(* IEC 61131-3 sources: JingjiangMoonbox/Application/Application/数据类型/通讯协议/月影, 10 files *)

(* ---- StParam_Mailbox.st ---- *)
(*@CES
Name=StParam_Mailbox
Type=Gvl
TypeGuid=2db5746d-d284-4425-9f7f-2663a34b0ebc
Guid=28298cb9-a045-46a0-b057-5251b4c14df2
HasDeclaration=True
HasImplementation=False
*)
{DECLARATION}
{attribute 'pack_mode' := '1'}
TYPE StParam_Mailbox :
STRUCT
	dwSemaphore						:DWORD;(*通讯旗语						*)
	dwPlateAdjustmentProf			:DWORD;(*纵向版快速调整量/bit24~bit31为请求信号/低24bit用来表示要调整的量<单位:0.01mm>/ 	*)
	iRapidAdjProf_h					:INT  ;(*横向快速对版量描述				*)
	iGateSa							:INT  ;(*第一波门位置					*)
	iGateSaEx						:INT  ;(*第二波门位置					*)
	rAdjust_V						:REAL ;(*纵向版修正量					*)
	rAdjust_H						:REAL ;(*横向版修正量					*)
	dwFlag_Ctl						:DWORD;(*套色控制标志					*)
	dwFlag_Sts						:DWORD;(*套色状态标志					*)
	wButtonFun_Lamp					:WORD ;(*HMI界面按钮及指示灯			*)
	wSwitchFun						:WORD ;(*界面开关*)
	wRsv							:WORD;
//2025.11.7.142851先把数据统一了，dwSlaveBtn_HMI分两个word,一个暂时baoliu
//	dwSlaveBtn_HMI					:DWORD;(*界面按钮						*)
	rStep_Pressure_Prn_Net			:REAL ;(*版辊网辊按钮步进量				*)
	rLong_Step_Roller_Pressure		:REAL ;(*色组压力控制长步进值			*)
	rShort_Step_Roller_Pressure		:REAL ;(*色组压力控制短步进值			*)
	wAirInletWindDoorValue			:WORD ;(*进风口风门开度值				*)
	wAirExhaustWindDoorValue		:WORD ;(*排风口风门开度值				*)
	wAirReturnWindDoorValue			:WORD ;(*回风口风门开度值				*)
	dwCtlBits_UnitBaseCraft			:DWORD;(*界面工艺开关及状态				*)
	wHz_UnitInkRoller_ManuallySet	:WORD ;(*递墨辊手动频率					*)
	wCoeff_UnitInkRoller_Auto		:WORD ;(*递墨辊自动系数					*)
	wHz_UnitScraper_ManuallySet		:WORD ;(*刮刀手动频率					*)
	wCoeff_UnitScraper_Auto			:WORD ;(*刮刀自动系数					*)
	wHz_UnitHotWind					:WORD ;(*热风频率						*)
	wHz_UnitHotWind_2				:WORD ;(*热风2频率						*)
	wSV_UnitTemCtl					:WORD ;(*加热设定温度					*)
	wUnit_output_I					:WORD ;(*IO监控输出1					*)
	wUnit_output_II					:WORD ;(*IO监控输出2					*)
	//xi.hy//新增
	bySignalSelect					:BYTE; (*光纤电眼信号选择*)
	rOffset_T1						:REAL;	//T1路光纤偏移
	rSource_Light_T1       			:REAL;  //T1路光纤光源
	rBias_T1			  			:REAL;  //T1路光纤电眼偏置
	rBrightness_Light_T1			:REAL;  //T1路光纤电眼亮度

	rOffset_T2						:REAL;  //T2路光纤偏移
	rSource_Light_T2				:REAL;  //T2路光纤光源
	rBias_T2						:REAL;  //T2路光纤电眼偏置
	rBrightness_Light_T2			:REAL;  //T2路光纤电眼亮度

	(*2025.8.14.143359增加一些参数*)
// 	wAccButton_Count				: WORD;
// 	wDecButton_Count			: WORD;
// 	wUpAdjButton_Count			: WORD;
// 	wDnAdjButton_Count			: WORD;
// 	wLeftAdjButton_Count			: WORD;
// 	wRightAdjButton_Count			: WORD;
// 	wAlarmButton_Count			: WORD;

	rHz_AxisAirBlowning_ManuallySet			: REAL;
	rHz_AxisAirExhaust_ManuallySet		: REAL;

	wSlaveBtn_HMI		: WORD;    //.0 版辊操作侧靠近
								   //.1 版辊操作侧远离
								   //.2 版辊平行靠近
								   //.3 版辊平行远离
								   //.4 版辊传动侧靠近
								   //.5 版辊传动侧远离
								   //.6 网辊操作侧靠近
								   //.7 网辊操作侧远离
								   //.8 网辊平行靠近
								   //.9 网辊平行远离
								   //.10 网辊传动侧靠近
								   //.11 网辊传动侧远离
								   //.12 版辊标定
								   //.13 网辊标定
								   //.14 张带棍标定
							 	   //.15 版辊合压
	wSlaveBtn_HMI2		: WORD;
									//. 0  版辊离压
									//. 1 网辊合压
									//. 2 网辊离压
									//. 3 版辊换版
									//. 4 网辊换版
									//. 5 自动换版
									//. 6 换版完成
									// .7 显示换版状态
	wButtonAndSwitch_ChaoXu	: WORD;	//.0 匀墨
										//.1 网辊锁轴
										//.2 充气
										//.3 墨盘电磁阀升
										//.4 照明
										//.5 显示是否修改版周
										//.6 确认修改版周
										//.7
										//.8
										//.9 版辊单动
										//.10 底辊单动
										//.11 合压
										//.12 离压
										//.13 横向左移
										//.14 横向右移

	uiRsv_data					: UINT;//压力电机步进量2026.02.07.143804
	iStep_Horz_Use						: INT;

	//xi.hy
	wState_FiberMove:WORD;	//光纤行走状态
						//.0 行走电机运动中
						//.1 基准色位置确认
						//.2 手动左移
						//.3 手动右移
						//.4 定长运动启动使能
						//.5 回零正限位触发
						//.6 宽度计算成功标志
						//.7 电机读取回来的限位信号
						//.8 基准位置同步完成
						//.9 基准位置同步中
						//.10 从站计算宽度使能
						//.11
						//.12
						//.13
						//.14
						//.15
	wAlarm_FiberMove:WORD;		//光纤行走报警
	iFiberMoveDistanceIn:INT;	//光纤行走距离输入 *10
	iPosCur_FiberMove:INT;		//光纤行走当前位置*10
	iWidth_FindMarkCenter:INT;	//光纤行走 计算出来的宽度*100
	//2026.5.9.182337
	//2026.04.28.132649 xi.hy新增@七号开始
	iStsSlave_FiberMove:INT;  // 光纤行走 从站运动状态机
	//2026.05.28.181612
	iFiberMoveBasePosFromSlave:INT;//基准位置@来自从站

END_STRUCT
END_TYPE

{IMPLEMENTATION}

(* ---- StParam_PDU_Dn.st ---- *)
(*@CES
Name=StParam_PDU_Dn
Type=Gvl
TypeGuid=2db5746d-d284-4425-9f7f-2663a34b0ebc
Guid=7cc610ea-6431-4c4c-b72a-07e9312a874d
HasDeclaration=True
HasImplementation=False
*)
{DECLARATION}
{attribute 'pack_mode' := '1'}
TYPE StParam_PDU_Dn :
STRUCT
	byPkgId						: BYTE;(*数据包ID*)
	abyPayLoad					: ARRAY [1..57] OF BYTE;(*数据可变区域*)
	wCHK						: WORD;(*校验码*)
END_STRUCT
END_TYPE

{IMPLEMENTATION}

(* ---- StParam_PDU_Up.st ---- *)
(*@CES
Name=StParam_PDU_Up
Type=Gvl
TypeGuid=2db5746d-d284-4425-9f7f-2663a34b0ebc
Guid=86ab3953-ed0c-4c63-9744-6672adabd60d
HasDeclaration=True
HasImplementation=False
*)
{DECLARATION}
{attribute 'pack_mode' := '1'}
TYPE StParam_PDU_Up :
STRUCT
	byPkgId						: BYTE;(*数据包ID*)
	abyPayLoad					: ARRAY [1..45] OF BYTE;(*数据可变区域*)
	wCHK						: WORD;(*校验码*)
	byIDX_V						: BYTE;(*纵向误差索引*)
	byIDX_H						: BYTE;(* 横向误差索引 *)
	iErr_V_Raw					: INT;(*纵向误差原始值-跟前色*)
	iErr_H_Raw					: INT;(*横向误差原始值-跟前色*)
	iErr_V_Raw_1				: INT;(*纵向误差原始值-跟任意色*)
	iErr_H_Raw_1				: INT;(*横向误差原始值-跟任意色*)
	uiFSampleCounter			: UINT;(*精采样计数*)
END_STRUCT
END_TYPE

{IMPLEMENTATION}

(* ---- StPdu_Dn_91.st ---- *)
(*@CES
Name=StPdu_Dn_91
Type=Gvl
TypeGuid=2db5746d-d284-4425-9f7f-2663a34b0ebc
Guid=22e1e21e-e973-4286-a59d-d3b41682a852
HasDeclaration=True
HasImplementation=False
*)
{DECLARATION}
{attribute 'pack_mode' := '1'}
TYPE StPdu_Dn_91 :
STRUCT
	byUnitId					:BYTE  ;(*机组号+系ID(最高位为系ID)*)
	rGirth_Sam					:REAL  ;(*采样版周长*)
	uiNum_Sam					:WORD  ;(*采样减速比分子*)
	uiDen_Sam					:WORD  ;(*采样减速比分母*)
	byCurrUsrLevel				:BYTE  ;(*用户权限*)
	iCompanyId					:INT   ;(*用户编号*)
	byLanguageId				:BYTE  ;(*语言选择*)
	byMinutes_ScrAutoSleep		:BYTE  ;(*屏幕休眠时间*)
	wUnit_input_I				:WORD  ;(*色组IO输入1*)
	wUnit_input_II				:WORD  ;(*色组IO输入2*)
	wUnit_input_III				:WORD  ;(*色组IO输入3*)
	wVelocity					:WORD  ;(*主机速度，单位0.1m/min*)
	wVel_Axis					:WORD  ;(*轴速度，单位0.1m/min*)
//	wComplexBit					:WORD  ;(*复合控制位描述*)
	wAxis_RollerDn				:WORD  ;(*轴压辊状态(bit0-1U,bit15-16U)*)
	wAxis_Alarm_Prn				:WORD  ;(*色组版辊报警状态(bit0-1U,bit15-16U)*)
	dwAlarmCode					:DWORD ;(*轴报警码*)
	wComplexFlag_AxisInching	:WORD  ;(*所有轴的单运行状态*)
	wComplexFlag_Linkage		:WORD  ;(*所有轴的联动状态*)
	wComplexFlag_Estop			:DWORD ;(*所有轴的急停状态*)
	wHMI_SwitchSts				:WORD  ;(*色组人机界面开关状态*)
	wSts_HorzManuPreReg			:WORD  ;(*横向手动预套准状态*)
	iPos_HorzManuPreReg			:INT   ;(*横向手动预套准位置*)
(*2025.8.6.205703增加*)
	bySts_Flag					:BYTE;(*色组状态*)
(*	dwAxis_SkipTheHeader 		:DWORD;(*让料头标志*)*)
	bySts_Machine				:BYTE;
	(*
		bit0: 印刷标志
		bit1: 空转标志
		bit2:
	*)
	//2025.11.14.155203||把误差状态发到从站，用于从站人机屏保实现9-1=8；
	byErrSts_V					: BYTE;
//用两个预留放低通滤波频率2025.11.15.132130|niu.j|8-2=6
	//Filter原本的wRsv在这里改一下改为从站精采样数据低通滤波频率
	uilowpasscutoff_hz				:UINT;

	abyRsv_91					:ARRAY [1..6] OF BYTE  ;(*预留空间*)
END_STRUCT
END_TYPE

{IMPLEMENTATION}

(* ---- StPdu_Dn_92.st ---- *)
(*@CES
Name=StPdu_Dn_92
Type=Gvl
TypeGuid=2db5746d-d284-4425-9f7f-2663a34b0ebc
Guid=45573361-4128-408d-910f-d2643f065581
HasDeclaration=True
HasImplementation=False
*)
{DECLARATION}
{attribute 'pack_mode' := '1'}
TYPE StPdu_Dn_92 :
STRUCT
	iCurveViewMaxRange				:INT;(*误差曲线量程上限		*)
	bySignalGain					:BYTE;(*光电眼IO控制			*)
	byMarkTypeId					:BYTE;(*标记形式				*)
	byMarkArrangeModalId			:BYTE;(*标记排列形式			*)
	byFakeThreshold_V				:BYTE;(*纵向飞点阀值@丝			*)
	byFakeThreshold_H				:BYTE;(*横向飞点阀值@丝			*)
	rAlarm_V						:REAL;(*纵向报警值@mm			*)
	rAlarm_H						:REAL;(*横向报警值@mm			*)
	byAve_v_extra_V					:BYTE;(*套色误差显示平均次数	*)
	byAve_v_extra_H					:BYTE;(*套色误差显示平均次数	*)
(*	dwFlag_Sts						: DWORD;(* 状态标志 *)
(*												/bit0.纵向自动 *)
(*												/bit1.横向自动
												/bit9.双极性*)
(*												/ *)
*)
	iGateWidthPhy					: INT ;(*波门宽度				*)
	byTriangleMark_SideC			: BYTE;(*梯形标记三角形纵向边长	*)
	byTriangleMark_SideB			: BYTE;(*梯形标记三角形横向边长	*)
	bySysSamplePrecision			: BYTE;(*系统采样精度			*)
	byArcFineSampleType				: BYTE;(*套色采样方式			*)
	iSampleCfgParam_ctl				: INT ;(*采样控制参数里的ctl		*)
	byColorIdCurrent				: BYTE;(*当前色序				*)
	byColorIdFollow					: BYTE;(*跟踪色序				*)
	abyColorIdList					: ARRAY [1..16] OF BYTE;(*色序列表				*)
	//bySignalSelect					:BYTE;(*光纤电眼信号选择		*)
	xEnable_Arc						: BOOL;(*套印使能开关			*)
	uiSource_Light_T1_Cur			: UINT;
	uiSource_Light_T2_Cur			: UINT;

	//xi.hy2026.5.9.104409
	wDirAndMode_FiberMove			:WORD;//光纤行走的方向和模式:低位方向,高位模式：0不运动 1连续运动 2定长运动 3回零运动
	uiVel_FiberMove					:UINT;//光纤行走的速度:mm/s *10
	uiDistanceOut_FiberMove			:UINT;//光纤行走的输出距离:mm *10
	uiPulsePerCycle_FiberMove		:UINT;//光纤行走的单圈脉冲:pluse

	abyRsv_92						: ARRAY [1..1] OF BYTE;(*套色参数预留			*)
END_STRUCT
END_TYPE

{IMPLEMENTATION}

(* ---- StPdu_Dn_93.st ---- *)
(*@CES
Name=StPdu_Dn_93
Type=Gvl
TypeGuid=2db5746d-d284-4425-9f7f-2663a34b0ebc
Guid=1bb7fc47-9e93-466c-a1c5-84993bb7c104
HasDeclaration=True
HasImplementation=False
*)
{DECLARATION}
{attribute 'pack_mode' := '1'}
TYPE StPdu_Dn_93 :
STRUCT
	dwControlComplexBits		:DWORD;(*开关状态			*)
	wHz_UnitInkRoller_CurrWR	:WORD ;(*递墨辊最终写入频率	*)
	wHz_UnitScraper_CurrWR		:WORD ;(*刮刀写入频率		*)
	wHz_UnitHotWind_CurrWR		:WORD ;(*热风写入频率		*)
	wHz_UnitHotWind2_CurrWR		:WORD ;(*热风2写入频率		*)
	rPV_UnitTemCtl				:REAL ;(*当前温度			*)
	wSTS_UnitTemCtl				:WORD ;(*温控状态			*)
(*2025.8.6.212214增加*)
	wHotWind_Print				:WORD;(*热风打开色组号*)
	byDriverType_Hor			:BYTE;(*横向的驱动器类型*)
	wPulseCtlInf  				:WORD;(*脉冲控制信息*)
	wPulse_1r					:WORD;(*1圈的脉冲数*)
	byPulseCtl_DisPerPulse 		:BYTE;(*单位脉冲距离*)
	byPulseCtlBit 				:BYTE;(*脉冲控制位*)

	//2026.1.24.193136增加色组监控信息下发niu.j||扭矩监控总共14字节|30-14=16
	iTorque_PrnRoller			: INT;//色组版辊扭矩|%/Nm。实际扭矩*10，保留一位小鼠
	iTorque_NetRoller			: INT;//色组网辊扭矩|%/Nm。实际扭矩*10，保留一位小鼠
	iTorque_BottomRoller		: INT;//色组底辊扭矩|%/Nm。实际扭矩*10，保留一位小鼠
	iTorque_Prn_PressRoller_M	: INT;//色组版辊压力操作侧扭矩|%/Nm。实际扭矩*10，保留一位小鼠
	iTorque_Prn_PressRoller_G	: INT;//色组版辊压力传动侧扭矩|%/Nm。实际扭矩*10，保留一位小鼠
	iTorque_Net_PressRoller_M	: INT;//色组网辊压力操作侧扭矩|%/Nm。实际扭矩*10，保留一位小鼠
	iTorque_Net_PressRoller_G	: INT;//色组网辊压力传动侧扭矩|%/Nm。实际扭矩*10，保留一位小鼠

	iVel_PrnRoller				: INT;//版辊速度
	iVel_BottomRoller			: INT;//底辊速度
	//2026.02.07.141032增加两个字节12-2
	iVel_NetRoller				: INT;//转速
	//2026.5.9.104649
	uiDistancePerCycle_FiberMove	:UINT;//光纤行走的单圈距离:mm *100

	abyRsv_93					:ARRAY [1..8] OF BYTE ;(*工艺参数预留		*)
	//2026.03.18.152620 |uiDistancePerCycle_FiberMove->uiDistancePerCycle_FiberMove|10->8

END_STRUCT
END_TYPE

{IMPLEMENTATION}

(* ---- StPdu_Dn_94.st ---- *)
(*@CES
Name=StPdu_Dn_94
Type=Gvl
TypeGuid=2db5746d-d284-4425-9f7f-2663a34b0ebc
Guid=4d2a344d-885f-40aa-a7e4-6cbaf8202632
HasDeclaration=True
HasImplementation=False
*)
{DECLARATION}
{attribute 'pack_mode' := '1'}
TYPE StPdu_Dn_94 :
STRUCT
	rPos_M_Prn_HandWheelCtl		:REAL;(*版辊压力操作侧位置-手轮显示						*)
	rPos_G_Prn_HandWheelCtl		:REAL;(*版辊压力传动侧位置-手轮显示						*)
	rPos_M_Net_HandWheelCtl		:REAL;(*网辊压力操作侧位置-手轮显示						*)
	rPos_G_Net_HandWheelCtl		:REAL;(*网辊压力传动侧位置-手轮显示						*)
	rPos_PrnRoller_Pressure_M	:REAL;(*版辊压力操作侧实时位置							*)
	rPos_PrnRoller_Pressure_G	:REAL;(*版辊压力传动侧实时位置							*)
	rPos_NetRoller_Pressure_M	:REAL;(*网辊压力操作侧实时位置							*)
	rPos_NetRoller_Pressure_G	:REAL;(*网辊压力传动侧实时位置							*)
	byCtlId_HandWheel			:BYTE;(*手轮控制ID										*)
	byCtlSts_HandWheel			:BYTE;(*手轮控制状态									*)
	wAxis_Alarm_Net				:WORD;(*色组网辊报警状态(bit0-1U,bit15-16U)				*)
	wAxis_Alarm_Bottom			:WORD;(*色组底辊报警状态(bit0-1U,bit15-16U)				*)
	wAxis_Alarm_Prn_M			:WORD;(*色组版辊压力操作侧报警状态(bit0-1U,bit15-16U)	*)
	wAxis_Alarm_Prn_G			:WORD;(*色组版辊压力传动侧报警状态(bit0-1U,bit15-16U)	*)
	wAxis_Alarm_Net_M			:WORD;(*色组网辊压力操作侧报警状态(bit0-1U,bit15-16U)	*)
	wAxis_Alarm_Net_G			:WORD;(*色组网辊压力传动侧报警状态(bit0-1U,bit15-16U)	*)
	wAxis_Alarm_Other			:WORD;(*整机其他轴报警状态								*)
	abyRsv_93					:array [1..9] of BYTE;(*柔印参数预留									*)
END_STRUCT
END_TYPE

{IMPLEMENTATION}

(* ---- StPdu_Dn_95.st ---- *)
(*@CES
Name=StPdu_Dn_95
Type=Gvl
TypeGuid=2db5746d-d284-4425-9f7f-2663a34b0ebc
Guid=8cf234ae-5b35-4b85-a488-2096eed3c062
HasDeclaration=True
HasImplementation=False
*)
{DECLARATION}
{attribute 'pack_mode' := '1'}
TYPE StPdu_Dn_95 :
STRUCT
	//全自动套印代码
	byWidth_Mark_Max						: BYTE;(*单个色标最大宽度-0.1mm*)
	byWidth_Mark_Min						: BYTE;(*单个色标最小宽度-0.1mm*)
	byMaxGap								: BYTE;(*最大间隙，-0.1mm*)
	bySimilarityThreshold					: BYTE;(*相似度阈值40%-70%,*)
	bySpotWidth								: BYTE;(*光斑宽度*10*)

	byFlag_CommFromMaster					: BYTE;(*	bit0: xFlag_AutoAdj_En; bit1: xFlag_FindFirstMark; bit2: xCurManuAdjust
														bit3:xFlag_FindPreMark  bit4:xPreCurManuAdjust ;bit5xFlag_GateMoveFinish*)
// 	iKcode_Mark_Interval					: INT;(*1色Kcode标与色标间隔- 单位 0.1mm*)
// 	iTaps_Mark_Interval						: INT;(*2色Taps标与色标间隔-单位0.1mm*)

	byMeanOffset							: BYTE; (*均值偏移 越大越找不到小色标，太小会出现较多信号导致直接失败*)
//2026.4.30.161528增加波形美化使能|占用5字节\|46-5=41
	xRsMorphFilter 								: BOOL;//美化标志
	abyRsMorphFilter_Rsv						: ARRAY [1..4] OF BYTE;
	//全自动套印下发模版
	aiCurModeMidPoint: ARRAY [1..4] OF INT;//当前色模版中心
	abyCurModeRadius:ARRAY [1..4] OF BYTE;//当前色模版半径
	aiPreModeMidPoint: ARRAY [1..4] OF INT;//前一色模版中心
	abyPreModeRadius:ARRAY [1..4] OF BYTE;//前一色模版半径
	byOuterCoff :BYTE ;//外滑窗系数 *10
	byInnerCoff	:BYTE;	//内滑窗系数 *10
	abyRsv_95		: ARRAY [1..19] OF BYTE;
	//2026.05.08.111411 屏蔽 iKcode_Mark_Interval iTaps_Mark_Interval 添加 aiCurModeMidPoint-> byInnerCoff 41+4-26=19
	//2026.4.30.161528 xRsMorphFilter->abyRsMorphFilter_Rsv |46-5=41

	//2026.03.17.133427 byWidth_Mark_Max->byMeanOffset 57-11=46
END_STRUCT
END_TYPE

{IMPLEMENTATION}

(* ---- StPdu_Up_05.st ---- *)
(*@CES
Name=StPdu_Up_05
Type=Gvl
TypeGuid=2db5746d-d284-4425-9f7f-2663a34b0ebc
Guid=a7996cd8-0fa8-4259-90b6-cff49420832c
HasDeclaration=True
HasImplementation=False
*)
{DECLARATION}
{attribute 'pack_mode' := '1'}
TYPE StPdu_Up_05 :
STRUCT
	dwSlaveVer					:DWORD;(*从站程序版本	*)
	wHz_UnitInkRoller_CurrrRD	:WORD ;(*读取的递墨辊频率*)
	wSts_UnitInkRoller			:WORD ;(*读取的递墨辊状态*)
	wHz_UnitScraper_CurrRD		:WORD ;(*读取的刮刀频率	*)
	wSTS_UnitScraper			:WORD ;(*读取的递墨辊状态*)
	wHz_UnitHotWind_CurrRD		:WORD ;(*读取的热风频率	*)
	wSTS_UnitHotWind			:WORD ;(*读取的热风状态	*)
	wHz_UnitHotWind2_CurrRD		:WORD ;(*读取的热风2频率	*)
	wSTS_UnitHotWind_2			:WORD ;(*读取的热风2状态	*)
	byCnt_Comm					:BYTE ;(*ARM通讯计数		*)
	(*2025.8.6.212503增加*)
	iEncValue_Hor				:INT;(*横向编码器值*)
	byStsBit2					:BYTE;(*状态位*)
	wPulse_Rd					:WORD;(*输出的脉冲数*)
	byStsBit					:BYTE;(*油墨槽状态*)

	iResult_VFollowpre_1stDerivate	: INT;(*YZJ计算误差*)(*18-2=16*)
	//2025.11.13.105908||上传基线和峰值16-8=8
	uiPeakValue_t1				: UINT;
	uiPeakValue_t2				: UINT;
	uiBaseUse_t1				: UINT;
	uiBaseUse_t2				: UINT;

	//全自动套印，已经用完了8个预留 8-8=0
	iCurLabelPos :INT;(*本色三角标位置，点数*)
	iPreLabelPos :INT;(*前色三角标位置，点数*)
	byFlag_CommFromSlave					: BYTE;(*bit0 xFlag_FindFirstSuccess 当前色成功找到 ;
													bit1 xFlag_FindPreSuccess 前一色成功找到
													bit2 当前色寻找完成
													bit3 精采样宽度计算完成
													bit4 从站全自动套印空闲中
													bit5 从站触发找本色
													bit6 从站触发找混色*)

	byDetectedSignalCount : BYTE;(*当前检测到色标个数*)
	byMarkStep:BYTE;(*当前全自动套印步骤*)
	byWidthRS :BYTE;//粗采样计算色标宽度 0.1mm

	//abyRsv_05					:ARRAY [1..8] OF BYTE ;(*参数预留		*)
END_STRUCT
END_TYPE

{IMPLEMENTATION}

(* ---- StUnitCmdQueue.st ---- *)
(*@CES
Name=StUnitCmdQueue
Type=Gvl
TypeGuid=2db5746d-d284-4425-9f7f-2663a34b0ebc
Guid=19a15640-4c7d-4711-b79a-2e35810a62a5
HasDeclaration=True
HasImplementation=False
*)
{DECLARATION}
{attribute 'pack_mode' := '1'}
TYPE StUnitCmdQueue :
STRUCT
	byCmdNum				: BYTE;(* 命令数量 *)
	byCmdIdx				: BYTE;(* 命令当前索引id *)
	aiCmdId					: ARRAY [1..MAX_CMD_NUM_PDU] OF INT;(* 命令id *)
END_STRUCT
END_TYPE

{IMPLEMENTATION}
